   #Core.Named := TRUE;
   #Core.RegIndex := 0;
   IF "FRK_Registry".Fault OR "FRK_Registry".Count < 0 OR "FRK_Registry".Count > 32
       OR #ParentIndex < 0 OR #ParentIndex > "FRK_Registry".Count OR #ParentIndex > 32 THEN
       "FRK_Registry".Fault := TRUE;
       RETURN;
   END_IF;
   IF #ParentIndex > 0 THEN
       IF NOT "FRK_Registry".Rows[#ParentIndex].Valid THEN
           "FRK_Registry".Fault := TRUE;
           RETURN;
       END_IF;
   END_IF;
   IF LEN(#InstancePath) > 254 THEN
       "FRK_Registry".Fault := TRUE;
       RETURN;
   END_IF;
   #Identity := WSTRING_TO_STRING(#InstancePath);
   #QuotePos := FIND(IN1 := #Identity, IN2 := '"');
   WHILE #QuotePos > 0 DO
       #Identity := DELETE(IN := #Identity, L := 1, P := #QuotePos);
       #QuotePos := FIND(IN1 := #Identity, IN2 := '"');
   END_WHILE;
   IF LEN(#Identity) > 80 OR LEN(#Identity) = 0 OR "FRK_Registry".Count >= 32 THEN
       "FRK_Registry".Fault := TRUE;
       RETURN;
   END_IF;
   "FRK_Registry".Count := "FRK_Registry".Count + 1;
   #RowIndex := "FRK_Registry".Count;
   #Core.RegIndex := #RowIndex;
   #Core.ParentIndex := #ParentIndex;
   #Core.ModuleType := #ModuleType;
   #Status.Name := #Identity;
   #Status.TypeKey := #TypeKey;
   #Status.ModuleType := #ModuleType;
   #Status.TileEnable := TRUE;
   "FRK_Registry".Rows[#RowIndex].Valid := TRUE;
   "FRK_Registry".Rows[#RowIndex].Parent := #ParentIndex;
   "FRK_Registry".Rows[#RowIndex].ModuleType := #ModuleType;
   "FRK_Registry".Rows[#RowIndex].TypeId := #TypeId;
   "FRK_Registry".Rows[#RowIndex].Capabilities := #Capabilities;
END_FUNCTION

FUNCTION "FRK_Sha256Pin" : Bool   // FC26, SCL
{ S7_Optimized_Access := 'TRUE' }
VERSION : 0.1
// Core section 7.7 prototype: volatile provider injection and independent root sessions.
//  User records are salted Core-compatible hashes, never commissioning plaintext.
// stored: AutoNumber true, IsIECCheckEnabled false, SetENOAutomatically false, UDAEnableTagReadback false
   VAR_INPUT
      Size : DInt;
   END_VAR
   VAR_IN_OUT
      Data : Array[0..47] of Byte;
      Digest : Array[0..31] of Byte;
   END_VAR
   VAR_TEMP
      BlockBytes : Array[0..63] of Byte;
      Words : Array[0..63] of DWord;
      Hash : Array[0..7] of DWord;
      Index : DInt;
      "A" : DWord;
      "B" : DWord;
      C : DWord;
      D : DWord;
      "E" : DWord;
      F : DWord;
      G : DWord;
      H : DWord;
      S0 : DWord;
      S1 : DWord;
      T1 : DWord;
      T2 : DWord;
      K : Array[0..63] of DWord;
   END_VAR
BEGIN

   #FRK_Sha256Pin := FALSE;
   #K[0] := DWORD#16#428A2F98;
   #K[1] := DWORD#16#71374491;
   #K[2] := DWORD#16#B5C0FBCF;
   #K[3] := DWORD#16#E9B5DBA5;
   #K[4] := DWORD#16#3956C25B;
   #K[5] := DWORD#16#59F111F1;
   #K[6] := DWORD#16#923F82A4;
   #K[7] := DWORD#16#AB1C5ED5;
   #K[8] := DWORD#16#D807AA98;
   #K[9] := DWORD#16#12835B01;
   #K[10] := DWORD#16#243185BE;
   #K[11] := DWORD#16#550C7DC3;
   #K[12] := DWORD#16#72BE5D74;
   #K[13] := DWORD#16#80DEB1FE;
   #K[14] := DWORD#16#9BDC06A7;
   #K[15] := DWORD#16#C19BF174;
   #K[16] := DWORD#16#E49B69C1;
   #K[17] := DWORD#16#EFBE4786;
   #K[18] := DWORD#16#0FC19DC6;
   #K[19] := DWORD#16#240CA1CC;
   #K[20] := DWORD#16#2DE92C6F;
   #K[21] := DWORD#16#4A7484AA;
   #K[22] := DWORD#16#5CB0A9DC;
   #K[23] := DWORD#16#76F988DA;
   #K[24] := DWORD#16#983E5152;
   #K[25] := DWORD#16#A831C66D;
   #K[26] := DWORD#16#B00327C8;
   #K[27] := DWORD#16#BF597FC7;
   #K[28] := DWORD#16#C6E00BF3;
   #K[29] := DWORD#16#D5A79147;
   #K[30] := DWORD#16#06CA6351;
   #K[31] := DWORD#16#14292967;
   #K[32] := DWORD#16#27B70A85;
   #K[33] := DWORD#16#2E1B2138;
   #K[34] := DWORD#16#4D2C6DFC;
   #K[35] := DWORD#16#53380D13;
   #K[36] := DWORD#16#650A7354;
   #K[37] := DWORD#16#766A0ABB;
   #K[38] := DWORD#16#81C2C92E;
   #K[39] := DWORD#16#92722C85;
   #K[40] := DWORD#16#A2BFE8A1;
   #K[41] := DWORD#16#A81A664B;
   #K[42] := DWORD#16#C24B8B70;
   #K[43] := DWORD#16#C76C51A3;
   #K[44] := DWORD#16#D192E819;
   #K[45] := DWORD#16#D6990624;
   #K[46] := DWORD#16#F40E3585;
   #K[47] := DWORD#16#106AA070;
   #K[48] := DWORD#16#19A4C116;
   #K[49] := DWORD#16#1E376C08;
   #K[50] := DWORD#16#2748774C;
   #K[51] := DWORD#16#34B0BCB5;
   #K[52] := DWORD#16#391C0CB3;
   #K[53] := DWORD#16#4ED8AA4A;
   #K[54] := DWORD#16#5B9CCA4F;
   #K[55] := DWORD#16#682E6FF3;
   #K[56] := DWORD#16#748F82EE;
   #K[57] := DWORD#16#78A5636F;
   #K[58] := DWORD#16#84C87814;
   #K[59] := DWORD#16#8CC70208;
   #K[60] := DWORD#16#90BEFFFA;
   #K[61] := DWORD#16#A4506CEB;
   #K[62] := DWORD#16#BEF9A3F7;
   #K[63] := DWORD#16#C67178F2;
   FOR #Index := 0 TO 31 DO
       #Digest[#Index] := 0;
   END_FOR;
   IF #Size < 0 OR #Size > 48 THEN
       RETURN;
   END_IF;
   // Authentication messages fit exactly one SHA-256 block.
   FOR #Index := 0 TO 63 DO
       #BlockBytes[#Index] := 0;
   END_FOR;
   FOR #Index := 0 TO #Size - 1 DO
       #BlockBytes[#Index] := #Data[#Index];
   END_FOR;
   #BlockBytes[#Size] := BYTE#16#80;
   #BlockBytes[62] := DWORD_TO_BYTE(SHR(IN := DINT_TO_DWORD(#Size * 8), N := 8));
   #BlockBytes[63] := DINT_TO_BYTE(#Size * 8);
   #Hash[0] := DWORD#16#6A09E667;
   #Hash[1] := DWORD#16#BB67AE85;
   #Hash[2] := DWORD#16#3C6EF372;
   #Hash[3] := DWORD#16#A54FF53A;
   #Hash[4] := DWORD#16#510E527F;
   #Hash[5] := DWORD#16#9B05688C;
   #Hash[6] := DWORD#16#1F83D9AB;
   #Hash[7] := DWORD#16#5BE0CD19;
   FOR #Index := 0 TO 15 DO
       #Words[#Index] := SHL(IN := BYTE_TO_DWORD(#BlockBytes[4 * #Index]), N := 24)
       OR SHL(IN := BYTE_TO_DWORD(#BlockBytes[4 * #Index + 1]), N := 16)
       OR SHL(IN := BYTE_TO_DWORD(#BlockBytes[4 * #Index + 2]), N := 8)
       OR BYTE_TO_DWORD(#BlockBytes[4 * #Index + 3]);
   END_FOR;
   FOR #Index := 16 TO 63 DO
       #S0 := ROR(IN := #Words[#Index - 15], N := 7) XOR ROR(IN := #Words[#Index - 15], N := 18) XOR SHR(IN := #Words[#Index - 15], N := 3);
       #S1 := ROR(IN := #Words[#Index - 2], N := 17) XOR ROR(IN := #Words[#Index - 2], N := 19) XOR SHR(IN := #Words[#Index - 2], N := 10);
       #Words[#Index] := UDINT_TO_DWORD(ULINT_TO_UDINT(UDINT_TO_ULINT(DWORD_TO_UDINT(#Words[#Index - 16])) + UDINT_TO_ULINT(DWORD_TO_UDINT(#S0)) + UDINT_TO_ULINT(DWORD_TO_UDINT(#Words[#Index - 7])) + UDINT_TO_ULINT(DWORD_TO_UDINT(#S1))));
   END_FOR;
   #A := #Hash[0];
   #B := #Hash[1];
   #C := #Hash[2];
   #D := #Hash[3];
   #E := #Hash[4];
   #F := #Hash[5];
   #G := #Hash[6];
   #H := #Hash[7];
   FOR #Index := 0 TO 63 DO
       #S1 := ROR(IN := #E, N := 6) XOR ROR(IN := #E, N := 11) XOR ROR(IN := #E, N := 25);
       #T1 := UDINT_TO_DWORD(ULINT_TO_UDINT(UDINT_TO_ULINT(DWORD_TO_UDINT(#H)) + UDINT_TO_ULINT(DWORD_TO_UDINT(#S1)) + UDINT_TO_ULINT(DWORD_TO_UDINT((#E AND #F) XOR ((NOT #E) AND #G))) + UDINT_TO_ULINT(DWORD_TO_UDINT(#K[#Index])) + UDINT_TO_ULINT(DWORD_TO_UDINT(#Words[#Index]))));
       #S0 := ROR(IN := #A, N := 2) XOR ROR(IN := #A, N := 13) XOR ROR(IN := #A, N := 22);
       #T2 := UDINT_TO_DWORD(ULINT_TO_UDINT(UDINT_TO_ULINT(DWORD_TO_UDINT(#S0)) + UDINT_TO_ULINT(DWORD_TO_UDINT((#A AND #B) XOR (#A AND #C) XOR (#B AND #C)))));
       #H := #G;
       #G := #F;
       #F := #E;
       #E := UDINT_TO_DWORD(ULINT_TO_UDINT(UDINT_TO_ULINT(DWORD_TO_UDINT(#D)) + UDINT_TO_ULINT(DWORD_TO_UDINT(#T1))));
       #D := #C;
       #C := #B;
       #B := #A;
       #A := UDINT_TO_DWORD(ULINT_TO_UDINT(UDINT_TO_ULINT(DWORD_TO_UDINT(#T1)) + UDINT_TO_ULINT(DWORD_TO_UDINT(#T2))));
   END_FOR;
   #Words[0] := #A;
   #Words[1] := #B;
   #Words[2] := #C;
   #Words[3] := #D;
   #Words[4] := #E;
   #Words[5] := #F;
   #Words[6] := #G;
   #Words[7] := #H;
   FOR #Index := 0 TO 7 DO
       #Hash[#Index] := UDINT_TO_DWORD(ULINT_TO_UDINT(UDINT_TO_ULINT(DWORD_TO_UDINT(#Hash[#Index])) + UDINT_TO_ULINT(DWORD_TO_UDINT(#Words[#Index]))));
       #Digest[4 * #Index] := DWORD_TO_BYTE(SHR(IN := #Hash[#Index], N := 24));
       #Digest[4 * #Index + 1] := DWORD_TO_BYTE(SHR(IN := #Hash[#Index], N := 16));
       #Digest[4 * #Index + 2] := DWORD_TO_BYTE(SHR(IN := #Hash[#Index], N := 8));
       #Digest[4 * #Index + 3] := DWORD_TO_BYTE(#Hash[#Index]);
   END_FOR;
   FOR #Index := 0 TO 63 DO
       #BlockBytes[#Index] := 0;
       #Words[#Index] := 0;
   END_FOR;
   #FRK_Sha256Pin := TRUE;
END_FUNCTION

FUNCTION "FRK_Start" : Void   // FC14, SCL
{ S7_Optimized_Access := 'TRUE' }
VERSION : 0.1
// stored: AutoNumber true, IsIECCheckEnabled false, SetENOAutomatically false, UDAEnableTagReadback false
   VAR_INPUT
      Supported : Bool;
      Timeout : Time;
      Label : String;
   END_VAR
   VAR_IN_OUT
      Core : "FRK_Core";
      Status : "ST_ModuleStatus";
   END_VAR
BEGIN

   #Core.CommandLabel := #Label;
   IF NOT #Supported THEN
       "FRK_Fault"(Core := #Core,
                   Status := #Status,
                   ReasonCode := 2008,
                   Description := WSTRING#'fraktal.command.unsupported');
   ELSIF #Timeout <= T#0ms THEN
       "FRK_Fault"(Core := #Core,
                   Status := #Status,
                   ReasonCode := 2004,
                   Description := WSTRING#'fraktal.command.timeout.invalid');
   ELSE
       #Core.TimeoutMs := DINT_TO_UDINT(TIME_TO_DINT(#Timeout));
   END_IF;
END_FUNCTION

FUNCTION "FRK_SyncRegistry" : Void   // FC2, SCL
{ S7_Optimized_Access := 'TRUE' }
VERSION : 0.1
// stored: AutoNumber true, IsIECCheckEnabled false, SetENOAutomatically false, UDAEnableTagReadback false
   VAR_INPUT
      Index : DInt;
      Status : "ST_ModuleStatus";
   END_VAR
BEGIN

   // Nested checks precede array access; do not depend on short-circuit AND.
   IF #Index < 1 OR #Index > "FRK_Registry".Count OR #Index > 32 THEN
       "FRK_Registry".Fault := TRUE;
       RETURN;
   END_IF;
   IF NOT "FRK_Registry".Rows[#Index].Valid THEN
       "FRK_Registry".Fault := TRUE;
       RETURN;
   END_IF;
   "FRK_Registry".Rows[#Index].Exec := #Status.State;
   "FRK_Registry".Rows[#Index].ReasonCode := #Status.Diagnostic.ReasonCode;
   "FRK_Registry".Rows[#Index].Severity := #Status.Diagnostic.Severity;
END_FUNCTION

FUNCTION "FRK_UnitCascade" : Void   // FC58, SCL
{ S7_Optimized_Access := 'TRUE' }
VERSION : 0.1
// stored: AutoNumber true, IsIECCheckEnabled false, SetENOAutomatically false, UDAEnableTagReadback false
   VAR_INPUT
      ParentUnit : "FRK_Unit";
      Supported : Array[0..6] of Bool;
   END_VAR
   VAR_IN_OUT
      Core : "FRK_Core";
      Unit : "FRK_Unit";
      Status : "ST_ModuleStatus";
      Policy : Array[0..6] of "ST_ModePolicy";
      Access : "FRK_Access";
      History : Array[1..16] of "ST_Diagnostic";
      Head : Int;
   END_VAR
   VAR_TEMP
      Request : "ST_HmiRequest";
   END_VAR
BEGIN

   IF NOT #ParentUnit.CascadePending THEN
       RETURN;
   END_IF;
   IF #ParentUnit.CascadeKind = 6 OR #ParentUnit.CascadeKind = 9 THEN
       #Unit.FollowStart := FALSE;
       #Request.Kind := #ParentUnit.CascadeKind;
       "FRK_UnitOperation"(Core := #Core,
                           Unit := #Unit,
                           Status := #Status,
                           Policy := #Policy,
                           Access := #Access,
                           Supported := #Supported,
                           Request := #Request,
                           Response := "FRK_UnitScratch".Response,
                           Trusted := TRUE);
       RETURN;
   END_IF;
   #Request.Kind := 3;
   #Request.IntValue := #ParentUnit.CascadeMode;
   "FRK_UnitOperation"(Core := #Core,
                       Unit := #Unit,
                       Status := #Status,
                       Policy := #Policy,
                       Access := #Access,
                       Supported := #Supported,
                       Request := #Request,
                       Response := "FRK_UnitScratch".Response,
                       Trusted := TRUE);
   IF NOT "FRK_UnitScratch".Response.Accepted THEN
       #Unit.FollowStart := FALSE;
       #Request.Kind := 6;
       "FRK_UnitOperation"(Core := #Core,
                           Unit := #Unit,
                           Status := #Status,
                           Policy := #Policy,
                           Access := #Access,
                           Supported := #Supported,
                           Request := #Request,
                           Response := "FRK_UnitScratch".Response,
                           Trusted := TRUE);
       // Core names this event but has no assigned E_Reason ordinal yet.
       "FRK_HistoryEvent"(History := #History,
                          Head := #Head,
                          Reason := 2008,
                          Description := WSTRING#'std.event.childModeUnsupported',
                          SourcePath := STRING_TO_WSTRING(#Status.Name));
   ELSE
       #Unit.FollowStart := #ParentUnit.CascadeKind = 5;
   END_IF;
END_FUNCTION

FUNCTION "FRK_UnitConsume" : Void   // FC45, SCL
{ S7_Optimized_Access := 'TRUE' }
VERSION : 0.1
// stored: AutoNumber true, IsIECCheckEnabled false, SetENOAutomatically false, UDAEnableTagReadback false
   VAR_INPUT
      Supported : Array[0..6] of Bool;
   END_VAR
   VAR_IN_OUT
      Core : "FRK_Core";
      Unit : "FRK_Unit";
      Status : "ST_ModuleStatus";
      Policy : Array[0..6] of "ST_ModePolicy";
      Access : "FRK_Access";
      Response : "ST_HmiResponse";
   END_VAR
BEGIN

   IF NOT #Unit.RequestPending THEN
       RETURN;
   END_IF;
   // The generated typed ownership walk serves the static manifest after children.
   IF #Unit.Request.Kind = 23 THEN
       #Unit.Request.Secret := '';
       RETURN;
   END_IF;
   "FRK_UnitOperation"(Core := #Core,
                       Unit := #Unit,
                       Status := #Status,
                       Policy := #Policy,
                       Access := #Access,
                       Supported := #Supported,
                       Request := #Unit.Request,
                       Response := #Response,
                       Trusted := FALSE);
   #Unit.Request.Secret := '';
END_FUNCTION

FUNCTION "FRK_UnitFinish" : Void   // FC50, SCL
{ S7_Optimized_Access := 'TRUE' }
VERSION : 0.1
// stored: AutoNumber true, IsIECCheckEnabled false, SetENOAutomatically false, UDAEnableTagReadback false
   VAR_IN_OUT
      Core : "FRK_Core";
      Unit : "FRK_Unit";
      Response : "ST_HmiResponse";
      Status : "ST_ModuleStatus";
      Part : "ST_PartContext";
      History : Array[1..16] of "ST_Diagnostic";
      Head : Int;
   END_VAR
BEGIN

   IF #Core.Exec = 3 THEN
       IF NOT #Unit.EvReset THEN
           #Unit.FaultLatched := TRUE;
       END_IF;
       IF NOT #Unit.PrevError THEN
           "FRK_PartAborted"(Core := #Core,
                             Unit := #Unit,
                             Status := #Status,
                             Part := #Part,
                             History := #History,
                             Head := #Head);
       END_IF;
   END_IF;
   #Unit.PrevError := #Core.Exec = 3;
   IF #Core.Exec = 2 OR #Core.Exec = 4 THEN
       #Unit.RunReq := FALSE;
   END_IF;
   IF #Unit.Clearing AND #Core.Exec = 0 THEN
       IF "FRK_DescendantsReady"(OwnerIndex := #Core.RegIndex) THEN
           #Unit.Clearing := FALSE;
       END_IF;
   END_IF;
   #Unit.AbortReq := FALSE;
   #Unit.ReleaseChildren := FALSE;
   #Unit.EvReset := FALSE;
   IF #Unit.RequestPending THEN
       #Response.AckSequence := #Unit.SeenSequence;
       #Unit.RequestPending := FALSE;
   END_IF;
END_FUNCTION

FUNCTION "FRK_UnitFollow" : Void   // FC59, SCL
{ S7_Optimized_Access := 'TRUE' }
VERSION : 0.1
// stored: AutoNumber true, IsIECCheckEnabled false, SetENOAutomatically false, UDAEnableTagReadback false
   VAR_INPUT
      Supported : Array[0..6] of Bool;
   END_VAR
   VAR_IN_OUT
      Core : "FRK_Core";
      Unit : "FRK_Unit";
      Status : "ST_ModuleStatus";
      Policy : Array[0..6] of "ST_ModePolicy";
      Access : "FRK_Access";
   END_VAR
   VAR_TEMP
      Request : "ST_HmiRequest";
   END_VAR
BEGIN

   IF #Unit.FollowStart AND NOT #Unit.ModePending AND NOT #Unit.Clearing THEN
       #Unit.FollowStart := FALSE;
       #Request.Kind := 5;
       "FRK_UnitOperation"(Core := #Core,
                           Unit := #Unit,
                           Status := #Status,
                           Policy := #Policy,
                           Access := #Access,
                           Supported := #Supported,
                           Request := #Request,
                           Response := "FRK_UnitScratch".Response,
                           Trusted := TRUE);
   END_IF;
END_FUNCTION

FUNCTION "FRK_UnitMailbox" : Void   // FC44, SCL
{ S7_Optimized_Access := 'TRUE' }
VERSION : 0.1
// stored: AutoNumber true, IsIECCheckEnabled false, SetENOAutomatically false, UDAEnableTagReadback false
   VAR_INPUT
      Supported : Array[0..6] of Bool;
   END_VAR
   VAR_IN_OUT
      Core : "FRK_Core";
      Unit : "FRK_Unit";
      Status : "ST_ModuleStatus";
      Policy : Array[0..6] of "ST_ModePolicy";
      Access : "FRK_Access";
      Request : "ST_HmiRequest";
      Response : "ST_HmiResponse";
   END_VAR
   VAR_TEMP
      SequenceBefore : UDInt;
   END_VAR
BEGIN

   #SequenceBefore := #Request.Sequence;
   IF #SequenceBefore = 0 OR #SequenceBefore = #Unit.SeenSequence THEN
       RETURN;
   END_IF;
   #Unit.Request := #Request;
   IF #Request.Sequence <> #SequenceBefore THEN
       #Unit.Request.Secret := '';
       RETURN;
   END_IF;
   #Request.Secret := '';
   #Unit.RequestUser := #Access.CurrentUser;
   #Unit.SeenSequence := #SequenceBefore;
   #Unit.RequestPending := TRUE;
END_FUNCTION

FUNCTION "FRK_UnitMode" : Void   // FC46, SCL
{ S7_Optimized_Access := 'TRUE' }
VERSION : 0.1
// stored: AutoNumber true, IsIECCheckEnabled false, SetENOAutomatically false, UDAEnableTagReadback false
   VAR_IN_OUT
      Core : "FRK_Core";
      Unit : "FRK_Unit";
   END_VAR
BEGIN

   IF #Unit.ModePending THEN
       IF #Core.Exec = 1 THEN
           #Core.EvModeExit := TRUE;
           #Core.HookResult := 0;
       ELSIF #Core.Exec = 0 AND NOT #Unit.Clearing THEN
           #Unit.Mode := #Unit.RequestedMode;
           #Unit.ModePending := FALSE;
           #Unit.ExitFirst := FALSE;
           #Core.EvModeChanged := TRUE;
       ELSE
           #Unit.RunReq := FALSE;
       END_IF;
   END_IF;
END_FUNCTION

FUNCTION "FRK_UnitModeResolve" : Void   // FC47, SCL
{ S7_Optimized_Access := 'TRUE' }
VERSION : 0.1
// stored: AutoNumber true, IsIECCheckEnabled false, SetENOAutomatically false, UDAEnableTagReadback false
   VAR_INPUT
      Policy : Array[0..6] of "ST_ModePolicy";
      Timeout : Time;
   END_VAR
   VAR_IN_OUT
      Core : "FRK_Core";
      Unit : "FRK_Unit";
      Status : "ST_ModuleStatus";
   END_VAR
BEGIN

   IF #Unit.ModePending THEN
       IF #Timeout <= T#0ms OR "FRK_Elapsed"(NewMs := "FRK_Clock".NowMs, OldMs := #Unit.ModeSince) >= DINT_TO_UDINT(TIME_TO_DINT(#Timeout)) THEN
           "FRK_Fault"(Core := #Core,
                       Status := #Status,
                       ReasonCode := 2001,
                       Description := WSTRING#'std.error.hmiRequestRejected');
           #Unit.ModePending := FALSE;
           #Unit.FollowStart := FALSE;
           #Unit.ReleaseChildren := TRUE;
           #Unit.Clearing := TRUE;
       ELSIF #Core.EvModeExit THEN
           #Unit.ExitFirst := FALSE;
           IF #Policy[#Unit.Mode].Style = 0 THEN
               #Unit.StopReq := TRUE;
           ELSIF #Core.HookResult <= 0 THEN
               #Unit.AbortReq := TRUE;
               #Unit.ReleaseChildren := TRUE;
               #Unit.Clearing := TRUE;
           END_IF;
       END_IF;
   END_IF;
END_FUNCTION

FUNCTION "FRK_UnitOperation" : Void   // FC43, SCL
{ S7_Optimized_Access := 'TRUE' }
VERSION : 0.1
// stored: AutoNumber true, IsIECCheckEnabled false, SetENOAutomatically false, UDAEnableTagReadback false
   VAR_INPUT
      Supported : Array[0..6] of Bool;
      Request : "ST_HmiRequest";
      Trusted : Bool;
   END_VAR
   VAR_IN_OUT
      Core : "FRK_Core";
      Unit : "FRK_Unit";
      Status : "ST_ModuleStatus";
      Policy : Array[0..6] of "ST_ModePolicy";
      Access : "FRK_Access";
      Response : "ST_HmiResponse";
   END_VAR
   VAR_TEMP
      Gate : DInt;
      Desired : DInt;
      Query : Bool;
      Level : DInt;
   END_VAR
BEGIN

   #Response.Accepted := FALSE;
   #Response.Diagnostic := WSTRING#'';
   #Response.Report.Count := 0;
   #Response.Report.Released := TRUE;
   #Gate := -1;
   #Desired := -1;
   #Query := FALSE;
   CASE #Request.Kind OF
       5:
           #Gate := 5;
           #Desired := 0;
       6:
           #Gate := 5;
           #Desired := 1;
       3:
           #Gate := 4;
           #Desired := #Request.IntValue;
           IF #Desired = -1 THEN
               #Desired := -2;
           END_IF;
       9:
           #Gate := 7;
       11:
           #Gate := 2;
       24, 25:
           #Gate := 8;
       15:
           #Gate := 5;
           #Desired := 0;
           #Query := TRUE;
       16:
           #Gate := 2;
           #Query := TRUE;
       17:
           #Gate := #Request.IntValue;
           #Desired := -1;
           #Query := TRUE;
       ELSE
           #Gate := -1;
   END_CASE;
   IF #Gate <> -1 OR #Request.Kind = 17 THEN
       "FRK_UnitRelease"(Core := #Core,
                         Unit := #Unit,
                         Status := #Status,
                         Policy := #Policy,
                         Access := #Access,
                         Supported := #Supported,
                         Report := #Response.Report,
                         Gate := #Gate,
                         Desired := #Desired,
                         Trusted := #Trusted);
       IF #Query THEN
           #Response.Accepted := TRUE;
       ELSIF #Response.Report.Released THEN
           CASE #Request.Kind OF
               5:
                   #Unit.StopReq := FALSE;
                   #Unit.RunReq := TRUE;
                   #Response.Accepted := TRUE;
               6:
                   #Unit.StopReq := #Core.Exec = 1;
                   IF NOT #Unit.StopReq THEN
                       #Unit.RunReq := FALSE;
                   END_IF;
                   #Unit.FollowStart := FALSE;
                   #Response.Accepted := TRUE;
               3:
                   IF #Desired <> #Unit.Mode THEN
                       #Unit.ExitFirst := TRUE;
                       #Unit.ModeSince := "FRK_Clock".NowMs;
                       #Unit.RequestedMode := #Desired;
                       #Unit.ModePending := TRUE;
                       IF #Unit.Mode = 1 THEN
                           #Unit.ReleaseChildren := TRUE;
                           #Unit.Clearing := TRUE;
                       END_IF;
                   END_IF;
                   #Response.Accepted := TRUE;
               9:
                   #Unit.EvReset := TRUE;
                   #Unit.ModePending := FALSE;
                   #Unit.ExitFirst := FALSE;
                   #Unit.RunReq := FALSE;
                   #Unit.AbortReq := #Core.Exec = 1;
                   #Unit.StopReq := FALSE;
                   #Unit.FollowStart := FALSE;
                   #Unit.ReleaseChildren := TRUE;
                   #Unit.Clearing := TRUE;
                   #Unit.FaultLatched := FALSE;
                   IF #Core.Exec = 3 THEN
                       #Core.Armed := TRUE;
                   END_IF;
                   #Response.Accepted := TRUE;
               24:
                   #Level := -1;
                   IF #Request.TextValue = WSTRING#'0' THEN
                       #Level := 0;
                   ELSIF #Request.TextValue = WSTRING#'1' THEN
                       #Level := 1;
                   ELSIF #Request.TextValue = WSTRING#'2' THEN
                       #Level := 2;
                   ELSIF #Request.TextValue = WSTRING#'3' THEN
                       #Level := 3;
                   ELSIF #Request.TextValue = WSTRING#'4' THEN
                       #Level := 4;
                   END_IF;
                   IF #Request.IntValue >= 0 AND #Request.IntValue <= 11 AND #Level >= 0 THEN
                       IF #Request.IntValue <> 8 OR #Level <= #Access.CurrentLevel THEN
                           #Access.Policy.Required[#Request.IntValue] := #Level;
                           #Response.Accepted := TRUE;
                       END_IF;
                   END_IF;
               25:
                   IF #Request.DurationMs <= 604800000 THEN
                       #Access.Policy.SessionTimeout := DINT_TO_TIME(UDINT_TO_DINT(#Request.DurationMs));
                       #Response.Accepted := TRUE;
                   END_IF;
               ELSE
                   // Manual acceptance is resolved by the generated typed route.
                   #Response.Accepted := FALSE;
           END_CASE;
       END_IF;
   ELSE
       CASE #Request.Kind OF
           1:
               "FRK_AccessLogin"(Access := #Access,
                                 User := #Request.User,
                                 Secret := #Request.Secret,
                                 Sequence := #Request.Sequence);
               // Consumption is acknowledged now; correlated result is asynchronous.
               #Response.Accepted := TRUE;
           2:
               "FRK_AccessLogout"(Access := #Access);
               #Response.Accepted := TRUE;
           ELSE
               #Response.Diagnostic := WSTRING#'std.error.unsupportedHmiRequest';
       END_CASE;
   END_IF;
   IF #Response.Accepted AND NOT #Query THEN
       IF #Request.Kind = 5 OR #Request.Kind = 6 OR #Request.Kind = 3 OR #Request.Kind = 9 THEN
           #Unit.CascadePending := TRUE;
           #Unit.CascadeKind := #Request.Kind;
           #Unit.CascadeMode := #Unit.Mode;
           IF #Request.Kind = 3 THEN
               #Unit.CascadeMode := #Desired;
           END_IF;
       END_IF;
   END_IF;
   IF NOT #Response.Accepted AND #Request.Kind <> 11 THEN
       IF #Response.Diagnostic = WSTRING#'' THEN
           #Response.Diagnostic := WSTRING#'std.error.hmiRequestRejected';
       END_IF;
       IF #Response.Report.Released THEN
           "FRK_ReleaseReason"(Report := #Response.Report,
                               Description := #Response.Diagnostic,
                               Reason := 2002,
                               Path := STRING_TO_WSTRING(#Status.Name),
                               Kind := 4);
       END_IF;
   END_IF;
END_FUNCTION

FUNCTION "FRK_UnitPrepare" : Void   // FC34, SCL
{ S7_Optimized_Access := 'TRUE' }
VERSION : 0.1
// Shared Unit services v0.1: operation authority, mailbox, modes and local carrier.
// stored: AutoNumber true, IsIECCheckEnabled false, SetENOAutomatically false, UDAEnableTagReadback false
   VAR_INPUT
      Startup : Bool;
      InitialMode : DInt;
   END_VAR
   VAR_IN_OUT
      Core : "FRK_Core";
      Unit : "FRK_Unit";
      Policy : Array[0..6] of "ST_ModePolicy";
      Request : "ST_HmiRequest";
      Response : "ST_HmiResponse";
   END_VAR
   VAR_TEMP
      Index : DInt;
   END_VAR
BEGIN

   #Core.EvModeExit := FALSE;
   #Core.EvModeChanged := FALSE;
   IF NOT #Unit.Initialized THEN
       #Unit.Initialized := TRUE;
       #Unit.Permit := TRUE;
       FOR #Index := 0 TO 7 - 1 DO
           #Policy[#Index].Shield := 1;
           #Policy[#Index].Style := 1;
       END_FOR;
       #Policy[0].Style := 0;
       #Policy[2].Shield := 0;
       #Policy[1].Shield := 0;
       #Policy[3].Shield := 2;
       #Policy[4].Shield := 2;
       #Unit.Mode := #InitialMode;
   END_IF;
   IF #Startup THEN
       #Unit.EvReset := FALSE;
       #Unit.Mode := #InitialMode;
       #Unit.RunReq := FALSE;
       #Unit.AbortReq := #Core.Exec = 1;
       #Unit.StopReq := FALSE;
       #Unit.ModePending := FALSE;
       #Unit.FollowStart := FALSE;
       #Unit.CascadePending := FALSE;
       #Unit.ReleaseChildren := TRUE;
       #Unit.Clearing := TRUE;
       // Consume the restart boundary without executing a transported request.
       #Unit.SeenSequence := #Request.Sequence;
       #Unit.RequestPending := FALSE;
       #Request.Secret := '';
       #Response.Accepted := FALSE;
       #Response.Diagnostic := WSTRING#'std.error.hmiRequestRejected';
       #Response.AckSequence := #Unit.SeenSequence;
   END_IF;
   IF #Core.ReleasePending THEN
       #Unit.FollowStart := FALSE;
       // An incoming parent mode/reset operation is already queued for this scan.
       // Preserve its cascade while cancelling the old command.
       #Unit.RunReq := FALSE;
       #Unit.AbortReq := TRUE;
       #Unit.ReleaseChildren := TRUE;
       #Unit.Clearing := TRUE;
   END_IF;
END_FUNCTION

FUNCTION "FRK_UnitRelease" : Void   // FC53, SCL
{ S7_Optimized_Access := 'TRUE' }
VERSION : 0.1
// stored: AutoNumber true, IsIECCheckEnabled false, SetENOAutomatically false, UDAEnableTagReadback false
   VAR_INPUT
      Gate : DInt;
      Desired : DInt;
      Trusted : Bool;
      Core : "FRK_Core";
      Unit : "FRK_Unit";
      Status : "ST_ModuleStatus";
      Policy : Array[0..6] of "ST_ModePolicy";
      Access : "FRK_Access";
      Supported : Array[0..6] of Bool;
   END_VAR
   VAR_IN_OUT
      Report : "ST_ReleaseReport";
   END_VAR
BEGIN

   #Report.Count := 0;
   #Report.Released := TRUE;
   IF #Gate <> 5 AND #Gate <> 4
       AND #Gate <> 7 AND #Gate <> 2
       AND #Gate <> 8 THEN
       "FRK_ReleaseReason"(Report := #Report,
                           Description := WSTRING#'std.error.unsupportedHmiRequest',
                           Reason := 2008,
                           Path := STRING_TO_WSTRING(#Status.Name),
                           Kind := 4);
       RETURN;
   END_IF;
   IF NOT #Trusted THEN
       IF #Access.CurrentLevel < #Access.Policy.Required[#Gate] THEN
           "FRK_ReleaseReason"(Report := #Report,
                               Description := WSTRING#'std.release.insufficientAction',
                               Reason := 2002,
                               Path := STRING_TO_WSTRING(#Status.Name),
                               Kind := 1);
       END_IF;
   END_IF;
   CASE #Gate OF
       5:
           // Desired=0 is Start, Desired=1 is Stop. Generic action query is Stop.
           IF #Desired = 0 THEN
               IF #Unit.Mode = 1 OR #Unit.ModePending THEN
                   "FRK_ReleaseReason"(Report := #Report,
                                       Description := WSTRING#'std.error.unsupportedModeRequest',
                                       Reason := 2002,
                                       Path := STRING_TO_WSTRING(#Status.Name),
                                       Kind := 0);
               END_IF;
               IF #Core.Exec <> 0 OR #Unit.RunReq OR #Unit.Clearing OR #Unit.FaultLatched THEN
                   "FRK_ReleaseReason"(Report := #Report,
                                       Description := WSTRING#'std.error.hmiRequestRejected',
                                       Reason := 2011,
                                       Path := STRING_TO_WSTRING(#Status.Name),
                                       Kind := 4);
               END_IF;
               IF NOT #Unit.Permit THEN
                   "FRK_ReleaseReason"(Report := #Report,
                                       Description := #Unit.PermitDiag.Description,
                                       Reason := #Unit.PermitDiag.ReasonCode,
                                       Path := #Unit.PermitDiag.SourcePath,
                                       Kind := 3);
               END_IF;
           END_IF;
       4:
           IF #Unit.ModePending THEN
               "FRK_ReleaseReason"(Report := #Report,
                                   Description := WSTRING#'std.release.modeChangeAlreadyPending',
                                   Reason := 2011,
                                   Path := STRING_TO_WSTRING(#Status.Name),
                                   Kind := 0);
           END_IF;
           IF #Core.Exec = 1 AND #Unit.Mode <> 1 THEN
               IF #Policy[#Unit.Mode].Shield = 2 THEN
                   "FRK_ReleaseReason"(Report := #Report,
                                       Description := WSTRING#'std.release.modeSwitchBlockedWhileRunning',
                                       Reason := 2002,
                                       Path := STRING_TO_WSTRING(#Status.Name),
                                       Kind := 0);
               END_IF;
           END_IF;
           IF #Desired <> -1 THEN
               IF #Desired < 0 OR #Desired >= 7 THEN
                   "FRK_ReleaseReason"(Report := #Report,
                                       Description := WSTRING#'std.error.unsupportedModeRequest',
                                       Reason := 2008,
                                       Path := STRING_TO_WSTRING(#Status.Name),
                                       Kind := 0);
               ELSIF NOT #Supported[#Desired] THEN
                   "FRK_ReleaseReason"(Report := #Report,
                                       Description := WSTRING#'std.error.unsupportedModeRequest',
                                       Reason := 2008,
                                       Path := STRING_TO_WSTRING(#Status.Name),
                                       Kind := 0);
               END_IF;
           END_IF;
       7:
           // The complete alarm model is separate; this gate owns the current latch.
           IF NOT #Unit.FaultLatched AND #Core.Exec = 0 AND NOT #Unit.Clearing AND NOT #Unit.ModePending AND NOT #Unit.FollowStart THEN
               IF "FRK_DescendantsReady"(OwnerIndex := #Core.RegIndex) THEN
                   "FRK_ReleaseReason"(Report := #Report,
                                       Description := WSTRING#'std.release.noBlockingAlarm',
                                       Reason := 2011,
                                       Path := STRING_TO_WSTRING(#Status.Name),
                                       Kind := 4);
               END_IF;
           END_IF;
       2:
           "FRK_ManualCommon"(Core := #Core,
                              Unit := #Unit,
                              Status := #Status,
                              Report := #Report);
       ELSE
           RETURN;
   END_CASE;
END_FUNCTION

FUNCTION "FRK_UnitRunStart" : Void   // FC48, SCL
{ S7_Optimized_Access := 'TRUE' }
VERSION : 0.1
// stored: AutoNumber true, IsIECCheckEnabled false, SetENOAutomatically false, UDAEnableTagReadback false
   VAR_INPUT
      Timeout : Time;
      Label : String;
   END_VAR
   VAR_IN_OUT
      Core : "FRK_Core";
      Status : "ST_ModuleStatus";
   END_VAR
BEGIN

   "FRK_Start"(Core := #Core,
               Status := #Status,
               Supported := TRUE,
               Timeout := #Timeout,
               Label := #Label);
   // A continuous run ends at Stop. Bounded commands/steps own progress timeouts.
   #Core.TimeoutMs := 0;
END_FUNCTION

FUNCTION "FRK_UnitSetLocalCarrier" : Void   // FC35, SCL
{ S7_Optimized_Access := 'TRUE' }
VERSION : 0.1
// stored: AutoNumber true, IsIECCheckEnabled false, SetENOAutomatically false, UDAEnableTagReadback false
   VAR_INPUT
      Index : DInt;
   END_VAR
   VAR_IN_OUT
      Unit : "FRK_Unit";
   END_VAR
BEGIN

   #Unit.CarrierIndex := 0;
   IF #Index < 1 OR #Index > 32 THEN
       RETURN;
   END_IF;
   "FRK_Carriers".Slots[#Index].Enabled := TRUE;
   "FRK_Carriers".Slots[#Index].Kind := 2;
   #Unit.CarrierIndex := #Index;
END_FUNCTION

FUNCTION "FRK_UnitSetPermit" : Void   // FC41, SCL
{ S7_Optimized_Access := 'TRUE' }
VERSION : 0.1
// stored: AutoNumber true, IsIECCheckEnabled false, SetENOAutomatically false, UDAEnableTagReadback false
   VAR_INPUT
      Ok : Bool;
      Diag : "ST_Diagnostic";
   END_VAR
   VAR_IN_OUT
      Unit : "FRK_Unit";
   END_VAR
BEGIN

   #Unit.Permit := #Ok;
   #Unit.PermitDiag := #Diag;
END_FUNCTION

DATA_BLOCK "GDB_FraktalMain"   // DB13
VERSION : 0.1
// stored: AutoNumber true, DBAccessibleFromOPCUA true, DBAccessibleFromWebserver true, InstanceOfName FB_FraktalMain, InstanceOfType FB
"FB_FraktalMain"
BEGIN
END_DATA_BLOCK

DATA_BLOCK "StationA"   // DB11
VERSION : 0.1
// stored: AutoNumber true, DBAccessibleFromOPCUA true, DBAccessibleFromWebserver true, InstanceOfName FB_DeclarationUnit, InstanceOfType FB
"FB_DeclarationUnit"
BEGIN
END_DATA_BLOCK

DATA_BLOCK "StationB"   // DB12
VERSION : 0.1
// stored: AutoNumber true, DBAccessibleFromOPCUA true, DBAccessibleFromWebserver true, InstanceOfName FB_DeclarationUnit, InstanceOfType FB
"FB_DeclarationUnit"
BEGIN
END_DATA_BLOCK
